FUNCTION_BLOCK "Tgp_InstanceEffect"
{ S7_Optimized_Access := 'TRUE' }
VERSION : 0.1
VAR_INPUT
 Enable : Bool;
END_VAR
VAR_OUTPUT
 Active : Bool;
END_VAR
VAR
 RetainedMarker : Int := 17;
 Child : "Tgp_TemplateFB_LAD";
END_VAR
BEGIN
 #Active := #Enable;
END_FUNCTION_BLOCK
